TYPE
    TcoKukaKss_Config_v_9_3_x :
    STRUCT
        InfoTime : TIME := T#2S;
        ErrorTime : TIME := T#0S;
		
    END_STRUCT
END_TYPE

(* stored: Version 1.1.0.1, ProductVersion 3.1.4024.12
   DUT TcoKukaKss_Config_v_9_3_x: Id {b0e199fc-e14e-461a-8c58-7d7770f14dcd} *)
